(* IEC 61131-3 sources: Test002/ConveyorBelt/Network/Network0, 1 file *)

(* ---- ONE_Network0_Table.st ---- *)
#define OBJECTS_CONFIG

FUNCTION GLOBAL TAB ONE_Network0
-1$UINT, 0$UINT,
0$UINT, 0$UINT,

1$UDINT,
TO_UDINT(3838332719), "ConveyorBelt", 1$UINT, 0$UINT, 2$UINT,

_NO_ATTR, TO_UDINT(686365345), "CONVEYORBELT1",
_NO_ATTR, TO_UDINT(2984266523), "CONVEYORBELT2",

//Internal connections
0$UDINT,
0$UDINT,
0$UDINT,
0$UDINT,

//Initialization values
0$UDINT,
5$UDINT,
TO_UDINT(0), "TimeDelay", TO_UDINT(5000),//|Network0.ConveyorBelt1.TimeDelay;
TO_UDINT(0), "ConveyorbeltSteps", TO_UDINT(ConveyorBelt::Step01),//|Network0.ConveyorBelt1.ConveyorbeltSteps;
TO_UDINT(0), "Motor", TO_UDINT(0),//|Network0.ConveyorBelt1.Motor;
TO_UDINT(1), "TimeDelay", TO_UDINT(5000),//|Network0.ConveyorBelt2.TimeDelay;
TO_UDINT(1), "ConveyorbeltSteps", TO_UDINT(Step01),//|Network0.ConveyorBelt2.ConveyorbeltSteps;

//Symbolic initialization values
0$UDINT,
0$UDINT,

//Initialization of string values
0$UDINT,
0$UDINT,

//Configuration of tasks (RealTime, Cyclic, Background)
0$UDINT,
0$UDINT,

0$UDINT,
2$UDINT,
TO_UDINT(0), (10)$UDINT, 4194303$DINT, 	//CONVEYORBELT1
TO_UDINT(1), (10)$UDINT, 4194303$DINT, 	//CONVEYORBELT2

0$UDINT,
0$UDINT,

//External connections
0$UDINT,
8$UDINT,
TO_UDINT(0), "Motor", C_DIR, TO_UDINT(2056942671), "DM1611","Output1",
TO_UDINT(0), "Lichtschrank", C_DIR, TO_UDINT(2056942671), "DM1611","Input2",
TO_UDINT(0), "Start", C_DIR, TO_UDINT(2056942671), "DM1611","Input1",
TO_UDINT(0), "Cylinder", C_DIR, TO_UDINT(2056942671), "DM1611","Output2",
TO_UDINT(1), "Motor", C_DIR, TO_UDINT(2056942671), "DM1611","Output3",
TO_UDINT(1), "Lichtschrank", C_DIR, TO_UDINT(2056942671), "DM1611","Input3",
TO_UDINT(1), "Start", C_DIR, TO_UDINT(2056942671), "DM1611","Input2",
TO_UDINT(1), "Cylinder", C_DIR, TO_UDINT(2056942671), "DM1611","Output4",

//Magic internal connections
0$UDINT,
0$UDINT,

//Configuration of timeslots of tasks (RealTime, Cyclic)
#ifdef __LSLLDR_TIMESLOTS__
0$UDINT,
0$UDINT,

0$UDINT,
0$UDINT,

#endif //__LSLLDR_TIMESLOTS__

//MultiMaster connections
#ifdef __LSLLDR_MULTIMASTER__
0$UDINT,
0$UDINT,
#endif //__LSLLDR_MULTIMASTER__

//Configuration for task ID (RealTime, CyclicTime)
#ifdef __LSLLDR_TASKID__
"\\\\TASKS2  "
0$UDINT,
0$UDINT,

0$UDINT,
2$UDINT,
(0)$UDINT, 	//CONVEYORBELT1
(0)$UDINT, 	//CONVEYORBELT2

0$UDINT,
0$UDINT,

#endif //__LSLLDR_TASKID__

END_FUNCTION
